FUNCTION_BLOCK TIME_ADD (* Basic Function Block Type *)
  (* Standard: 61499-2 *)
  (* Version 0.0, 10/5/2026, Schneider Electric, Template *)
  PACKAGE SE.Nereda;
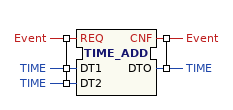
  EVENT_INPUT
    REQ WITH DT1, DT2; (* Normal Execution Request *)
  END_EVENT
  EVENT_OUTPUT
    CNF WITH DTO; (* Execution Confirmation *)
  END_EVENT
  VAR_INPUT
    DT1 : TIME; (* Input event qualifier *)
    DT2 : TIME;
  END_VAR
  VAR_OUTPUT
    DTO : TIME; (* Output event qualifier *)
  END_VAR
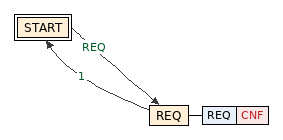
  EC_STATES
    START; (* Initial State *)
    REQ : REQ -> CNF; (* Normal execution *)
  END_STATES
  EC_TRANSITIONS
    START TO REQ := REQ;
    REQ TO START := 1;
  END_TRANSITIONS
  ALGORITHM REQ IN ST: (* Normally executed algorithm *)
;
DTO := DT1 + DT2;
  END_ALGORITHM
END_FUNCTION_BLOCK
